Universal Robots URScript: Jonathan_code.script

  # Default parameters:
  global speed_ms = 0.3
  global speed_rads = 0.75
  global accel_mss = 3
  global accel_radss = 1.2
  global blend_radius_m = 0.001

  # Add subprograms here
  # Start of main program
  # Program generated by RoboDK v5.6.5 for UR10e on 12/10/2023 11:38:14
  # Using nominal kinematics.
  blend_radius_m = 0.001
  speed_ms = 1.000
  # set_reference(p[0.335000, -0.154000, 0.000000, 0.000000, 0.000000, 0.000000])
  set_tcp(p[0.000000, 0.000000, 0.253000, 0.000000, 0.000000, 0.000000])
  # Show Tool
  movej([0.470150, -1.112535, -2.574781, -1.025073, 1.570796, 2.040947],accel_radss,speed_rads,0,blend_radius_m
  movel([0.470150, -1.206188, -2.638649, -0.867552, 1.570796, 2.040947],accel_mss,speed_ms,0,blend_radius_m)
  speed_ms = 1.000
  movel([0.470150, -1.233460, -2.652834, -0.826095, 1.570796, 2.040947],accel_mss,speed_ms,0,blend_radius_m)
  speed_ms = 0.003
  movel([0.470150, -1.244207, -2.658024, -0.810158, 1.570796, 2.040947],accel_mss,speed_ms,0,blend_radius_m)
  speed_ms = 0.007
  movel([0.482800, -1.244203, -2.658026, -0.810160, 1.570796, 2.053597],accel_mss,speed_ms,0,blend_radius_m)
  movel([0.495365, -1.244373, -2.657937, -0.810079, 1.570796, 2.066162],accel_mss,speed_ms,0,blend_radius_m)
  movel([0.493680, -1.247797, -2.656131, -0.808461, 1.570796, 2.064476],accel_mss,speed_ms,0,blend_radius_m)
  movel([0.492007, -1.251200, -2.654322, -0.806866, 1.570796, 2.062803],accel_mss,speed_ms,0,blend_radius_m)
  movel([0.479519, -1.251033, -2.654411, -0.806944, 1.570796, 2.050316],accel_mss,speed_ms,0,blend_radius_m)
  movel([0.466949, -1.251037, -2.654410, -0.806943, 1.570796, 2.037745],accel_mss,speed_ms,0,blend_radius_m)
  movel([0.468544, -1.247632, -2.656219, -0.808539, 1.570796, 2.039340],accel_mss,speed_ms,0,blend_radius_m)
  movel([0.470150, -1.244207, -2.658024, -0.810158, 1.570796, 2.040947],accel_mss,speed_ms,0,blend_radius_m)
  speed_ms = 0.003
  movel([0.470150, -1.247853, -2.659738, -0.804798, 1.570796, 2.040947],accel_mss,speed_ms,0,blend_radius_m)
  speed_ms = 0.007
  movel([0.482800, -1.247850, -2.659740, -0.804799, 1.570796, 2.053597],accel_mss,speed_ms,0,blend_radius_m)
  movel([0.495365, -1.248020, -2.659650, -0.804719, 1.570796, 2.066162],accel_mss,speed_ms,0,blend_radius_m)
  movel([0.493680, -1.251437, -2.657839, -0.803114, 1.570796, 2.064476],accel_mss,speed_ms,0,blend_radius_m)
  movel([0.492007, -1.254834, -2.656024, -0.801531, 1.570796, 2.062803],accel_mss,speed_ms,0,blend_radius_m)
  movel([0.479519, -1.254667, -2.656113, -0.801608, 1.570796, 2.050316],accel_mss,speed_ms,0,blend_radius_m)
  movel([0.466949, -1.254671, -2.656111, -0.801607, 1.570796, 2.037745],accel_mss,speed_ms,0,blend_radius_m)
  movel([0.468544, -1.251272, -2.657926, -0.803191, 1.570796, 2.039340],accel_mss,speed_ms,0,blend_radius_m)
  movel([0.470150, -1.247853, -2.659738, -0.804798, 1.570796, 2.040947],accel_mss,speed_ms,0,blend_radius_m)
  speed_ms = 0.003
  movel([0.470150, -1.233460, -2.652834, -0.826095, 1.570796, 2.040947],accel_mss,speed_ms,0,blend_radius_m)
  speed_ms = 1.000
  movel([0.470150, -1.206188, -2.638649, -0.867552, 1.570796, 2.040947],accel_mss,speed_ms,0,blend_radius_m)
  movel([0.500005, -1.181387, -2.650684, -0.880318, 1.570796, 2.070801],accel_mss,speed_ms,0,blend_radius_m)
  movel([0.500005, -1.208894, -2.665198, -0.838297, 1.570796, 2.070801],accel_mss,speed_ms,0,blend_radius_m)
  speed_ms = 0.003
  movel([0.500005, -1.219758, -2.670513, -0.822118, 1.570796, 2.070801],accel_mss,speed_ms,0,blend_radius_m)
  speed_ms = 0.007
  movel([0.496713, -1.215452, -2.672641, -0.824296, 1.570796, 2.067509],accel_mss,speed_ms,0,blend_radius_m)
  movel([0.497565, -1.208277, -2.676141, -0.827971, 1.570796, 2.068361],accel_mss,speed_ms,0,blend_radius_m)
  movel([0.502312, -1.200573, -2.679835, -0.831981, 1.570796, 2.073109],accel_mss,speed_ms,0,blend_radius_m)
  movel([0.509447, -1.194948, -2.682491, -0.834950, 1.570796, 2.080243],accel_mss,speed_ms,0,blend_radius_m)
  movel([0.511019, -1.194268, -2.682810, -0.835312, 1.570796, 2.081816],accel_mss,speed_ms,0,blend_radius_m)
  movel([0.512848, -1.193698, -2.683076, -0.835615, 1.570796, 2.083644],accel_mss,speed_ms,0,blend_radius_m)
  movel([0.514636, -1.193318, -2.683254, -0.835817, 1.570796, 2.085432],accel_mss,speed_ms,0,blend_radius_m)
  movel([0.516087, -1.193207, -2.683306, -0.835876, 1.570796, 2.086884],accel_mss,speed_ms,0,blend_radius_m)
  movel([0.521675, -1.195790, -2.682095, -0.834503, 1.570796, 2.092471],accel_mss,speed_ms,0,blend_radius_m)
  movel([0.522729, -1.202299, -2.679013, -0.831077, 1.570796, 2.093526],accel_mss,speed_ms,0,blend_radius_m)
  movel([0.518940, -1.210348, -2.675137, -0.826904, 1.570796, 2.089737],accel_mss,speed_ms,0,blend_radius_m)
  movel([0.511727, -1.217078, -2.671840, -0.823471, 1.570796, 2.082524],accel_mss,speed_ms,0,blend_radius_m)
  movel([0.508244, -1.219012, -2.670883, -0.822493, 1.570796, 2.079040],accel_mss,speed_ms,0,blend_radius_m)
  movel([0.505130, -1.220107, -2.670340, -0.821942, 1.570796, 2.075926],accel_mss,speed_ms,0,blend_radius_m)
  movel([0.502386, -1.220345, -2.670222, -0.821823, 1.570796, 2.073182],accel_mss,speed_ms,0,blend_radius_m)
  movel([0.500005, -1.219758, -2.670513, -0.822118, 1.570796, 2.070801],accel_mss,speed_ms,0,blend_radius_m)
  speed_ms = 0.003
  movel([0.500005, -1.223447, -2.672269, -0.816673, 1.570796, 2.070801],accel_mss,speed_ms,0,blend_radius_m)
  speed_ms = 0.007
  movel([0.496713, -1.219148, -2.674405, -0.818836, 1.570796, 2.067509],accel_mss,speed_ms,0,blend_radius_m)
  movel([0.497565, -1.211984, -2.677917, -0.822488, 1.570796, 2.068361],accel_mss,speed_ms,0,blend_radius_m)
  movel([0.502312, -1.204292, -2.681624, -0.826473, 1.570796, 2.073109],accel_mss,speed_ms,0,blend_radius_m)
  movel([0.509447, -1.198675, -2.684289, -0.829425, 1.570796, 2.080243],accel_mss,speed_ms,0,blend_radius_m)
  movel([0.511019, -1.197995, -2.684609, -0.829784, 1.570796, 2.081816],accel_mss,speed_ms,0,blend_radius_m)
  movel([0.512848, -1.197426, -2.684877, -0.830086, 1.570796, 2.083644],accel_mss,speed_ms,0,blend_radius_m)
  movel([0.514636, -1.197048, -2.685055, -0.830287, 1.570796, 2.085432],accel_mss,speed_ms,0,blend_radius_m)
  movel([0.516087, -1.196936, -2.685107, -0.830346, 1.570796, 2.086884],accel_mss,speed_ms,0,blend_radius_m)
  movel([0.521675, -1.199516, -2.683892, -0.828981, 1.570796, 2.092471],accel_mss,speed_ms,0,blend_radius_m)
  movel([0.522729, -1.206015, -2.680799, -0.825575, 1.570796, 2.093526],accel_mss,speed_ms,0,blend_radius_m)
  movel([0.518940, -1.214052, -2.676909, -0.821428, 1.570796, 2.089737],accel_mss,speed_ms,0,blend_radius_m)
  movel([0.511727, -1.220771, -2.673601, -0.818017, 1.570796, 2.082524],accel_mss,speed_ms,0,blend_radius_m)
  movel([0.508244, -1.222703, -2.672640, -0.817046, 1.570796, 2.079040],accel_mss,speed_ms,0,blend_radius_m)
  movel([0.505130, -1.223795, -2.672095, -0.816499, 1.570796, 2.075926],accel_mss,speed_ms,0,blend_radius_m)
  movel([0.502386, -1.224033, -2.671976, -0.816380, 1.570796, 2.073182],accel_mss,speed_ms,0,blend_radius_m)
  movel([0.500005, -1.223447, -2.672269, -0.816673, 1.570796, 2.070801],accel_mss,speed_ms,0,blend_radius_m)
  speed_ms = 0.003
  movel([0.500005, -1.208894, -2.665198, -0.838297, 1.570796, 2.070801],accel_mss,speed_ms,0,blend_radius_m)
  speed_ms = 1.000
  movel([0.500005, -1.181387, -2.650684, -0.880318, 1.570796, 2.070801],accel_mss,speed_ms,0,blend_radius_m)
  movel([0.502939, -1.178463, -2.652060, -0.881866, 1.570796, 2.073735],accel_mss,speed_ms,0,blend_radius_m)
  movel([0.502939, -1.205994, -2.666612, -0.839782, 1.570796, 2.073735],accel_mss,speed_ms,0,blend_radius_m)
  speed_ms = 0.003
  movel([0.502939, -1.216871, -2.671942, -0.823575, 1.570796, 2.073735],accel_mss,speed_ms,0,blend_radius_m)
  speed_ms = 0.007
  movel([0.501818, -1.216382, -2.672184, -0.823824, 1.570796, 2.072614],accel_mss,speed_ms,0,blend_radius_m)
  movel([0.500967, -1.215437, -2.672649, -0.824303, 1.570796, 2.071763],accel_mss,speed_ms,0,blend_radius_m)
  movel([0.500167, -1.213807, -2.673449, -0.825133, 1.570796, 2.070964],accel_mss,speed_ms,0,blend_radius_m)
  movel([0.499493, -1.211784, -2.674438, -0.826167, 1.570796, 2.070289],accel_mss,speed_ms,0,blend_radius_m)
  movel([0.499454, -1.210389, -2.675117, -0.826883, 1.570796, 2.070250],accel_mss,speed_ms,0,blend_radius_m)
  movel([0.499992, -1.208799, -2.675888, -0.827701, 1.570796, 2.070788],accel_mss,speed_ms,0,blend_radius_m)
  movel([0.501476, -1.206040, -2.677221, -0.829128, 1.570796, 2.072272],accel_mss,speed_ms,0,blend_radius_m)
  movel([0.504659, -1.201513, -2.679388, -0.831488, 1.570796, 2.075455],accel_mss,speed_ms,0,blend_radius_m)
  movel([0.508226, -1.198314, -2.680906, -0.833169, 1.570796, 2.079022],accel_mss,speed_ms,0,blend_radius_m)
  movel([0.512021, -1.196627, -2.681702, -0.834060, 1.570796, 2.082817],accel_mss,speed_ms,0,blend_radius_m)
  movel([0.515863, -1.196480, -2.681771, -0.834138, 1.570796, 2.086659],accel_mss,speed_ms,0,blend_radius_m)
  movel([0.517050, -1.196870, -2.681587, -0.833932, 1.570796, 2.087846],accel_mss,speed_ms,0,blend_radius_m)
  movel([0.518044, -1.197576, -2.681254, -0.833558, 1.570796, 2.088840],accel_mss,speed_ms,0,blend_radius_m)
  movel([0.518815, -1.198576, -2.680782, -0.833031, 1.570796, 2.089612],accel_mss,speed_ms,0,blend_radius_m)
  movel([0.519336, -1.199836, -2.680185, -0.832368, 1.570796, 2.090133],accel_mss,speed_ms,0,blend_radius_m)
  movel([0.518927, -1.205179, -2.677634, -0.829575, 1.570796, 2.089724],accel_mss,speed_ms,0,blend_radius_m)
  movel([0.515430, -1.211016, -2.674812, -0.826561, 1.570796, 2.086227],accel_mss,speed_ms,0,blend_radius_m)
  movel([0.510067, -1.215433, -2.672651, -0.824305, 1.570796, 2.080863],accel_mss,speed_ms,0,blend_radius_m)
  movel([0.504562, -1.217042, -2.671858, -0.823489, 1.570796, 2.075358],accel_mss,speed_ms,0,blend_radius_m)
  movel([0.502939, -1.216871, -2.671942, -0.823575, 1.570796, 2.073735],accel_mss,speed_ms,0,blend_radius_m)
  speed_ms = 0.003
  movel([0.502939, -1.220565, -2.673703, -0.818121, 1.570796, 2.073735],accel_mss,speed_ms,0,blend_radius_m)
  speed_ms = 0.007
  movel([0.501818, -1.220076, -2.673945, -0.818367, 1.570796, 2.072614],accel_mss,speed_ms,0,blend_radius_m)
  movel([0.500967, -1.219134, -2.674412, -0.818844, 1.570796, 2.071763],accel_mss,speed_ms,0,blend_radius_m)
  movel([0.500167, -1.217506, -2.675215, -0.819668, 1.570796, 2.070964],accel_mss,speed_ms,0,blend_radius_m)
  movel([0.499493, -1.215486, -2.676207, -0.820696, 1.570796, 2.070289],accel_mss,speed_ms,0,blend_radius_m)
  movel([0.499454, -1.214093, -2.676889, -0.821407, 1.570796, 2.070250],accel_mss,speed_ms,0,blend_radius_m)
  movel([0.499992, -1.212506, -2.677663, -0.822220, 1.570796, 2.070788],accel_mss,speed_ms,0,blend_radius_m)
  movel([0.501476, -1.209751, -2.679000, -0.823638, 1.570796, 2.072272],accel_mss,speed_ms,0,blend_radius_m)
  movel([0.504659, -1.205231, -2.681175, -0.825983, 1.570796, 2.075455],accel_mss,speed_ms,0,blend_radius_m)
  movel([0.508226, -1.202036, -2.682698, -0.827655, 1.570796, 2.079022],accel_mss,speed_ms,0,blend_radius_m)
  movel([0.512021, -1.200352, -2.683497, -0.828540, 1.570796, 2.082817],accel_mss,speed_ms,0,blend_radius_m)
  movel([0.515863, -1.200205, -2.683566, -0.828617, 1.570796, 2.086659],accel_mss,speed_ms,0,blend_radius_m)
  movel([0.517050, -1.200594, -2.683382, -0.828413, 1.570796, 2.087846],accel_mss,speed_ms,0,blend_radius_m)
  movel([0.518044, -1.201300, -2.683048, -0.828041, 1.570796, 2.088840],accel_mss,speed_ms,0,blend_radius_m)
  movel([0.518815, -1.202298, -2.682574, -0.827517, 1.570796, 2.089612],accel_mss,speed_ms,0,blend_radius_m)
  movel([0.519336, -1.203556, -2.681975, -0.826858, 1.570796, 2.090133],accel_mss,speed_ms,0,blend_radius_m)
  movel([0.518927, -1.208892, -2.679415, -0.824082, 1.570796, 2.089724],accel_mss,speed_ms,0,blend_radius_m)
  movel([0.515430, -1.214719, -2.676583, -0.821087, 1.570796, 2.086227],accel_mss,speed_ms,0,blend_radius_m)
  movel([0.510067, -1.219129, -2.674414, -0.818846, 1.570796, 2.080863],accel_mss,speed_ms,0,blend_radius_m)
  movel([0.504562, -1.220735, -2.673619, -0.818035, 1.570796, 2.075358],accel_mss,speed_ms,0,blend_radius_m)
  movel([0.502939, -1.220565, -2.673703, -0.818121, 1.570796, 2.073735],accel_mss,speed_ms,0,blend_radius_m)
  speed_ms = 0.003
  movel([0.502939, -1.205994, -2.666612, -0.839782, 1.570796, 2.073735],accel_mss,speed_ms,0,blend_radius_m)
  speed_ms = 1.000
  movel([0.502939, -1.178463, -2.652060, -0.881866, 1.570796, 2.073735],accel_mss,speed_ms,0,blend_radius_m)
  movel([0.506130, -1.175000, -2.653677, -0.883712, 1.570796, 2.076926],accel_mss,speed_ms,0,blend_radius_m)
  movel([0.506130, -1.202560, -2.668276, -0.841553, 1.570796, 2.076926],accel_mss,speed_ms,0,blend_radius_m)
  speed_ms = 0.003
  movel([0.506130, -1.213452, -2.673623, -0.825314, 1.570796, 2.076926],accel_mss,speed_ms,0,blend_radius_m)
  speed_ms = 0.007
  movel([0.503262, -1.211890, -2.674386, -0.826113, 1.570796, 2.074059],accel_mss,speed_ms,0,blend_radius_m)
  movel([0.503107, -1.207977, -2.676286, -0.828126, 1.570796, 2.073904],accel_mss,speed_ms,0,blend_radius_m)
  movel([0.505736, -1.203530, -2.678425, -0.830434, 1.570796, 2.076532],accel_mss,speed_ms,0,blend_radius_m)
  movel([0.509953, -1.200615, -2.679815, -0.831959, 1.570796, 2.080749],accel_mss,speed_ms,0,blend_radius_m)
  movel([0.512348, -1.199943, -2.680134, -0.832312, 1.570796, 2.083144],accel_mss,speed_ms,0,blend_radius_m)
  movel([0.514007, -1.199944, -2.680134, -0.832311, 1.570796, 2.084803],accel_mss,speed_ms,0,blend_radius_m)
  movel([0.515159, -1.200632, -2.679807, -0.831950, 1.570796, 2.085955],accel_mss,speed_ms,0,blend_radius_m)
  movel([0.515994, -1.202071, -2.679122, -0.831196, 1.570796, 2.086790],accel_mss,speed_ms,0,blend_radius_m)
  movel([0.515943, -1.205637, -2.677415, -0.829338, 1.570796, 2.086739],accel_mss,speed_ms,0,blend_radius_m)
  movel([0.513721, -1.209501, -2.675548, -0.827340, 1.570796, 2.084517],accel_mss,speed_ms,0,blend_radius_m)
  movel([0.510054, -1.212409, -2.674133, -0.825847, 1.570796, 2.080851],accel_mss,speed_ms,0,blend_radius_m)
  movel([0.506130, -1.213452, -2.673623, -0.825314, 1.570796, 2.076926],accel_mss,speed_ms,0,blend_radius_m)
  speed_ms = 0.003
  movel([0.506130, -1.217151, -2.675389, -0.819848, 1.570796, 2.076926],accel_mss,speed_ms,0,blend_radius_m)
  speed_ms = 0.007
  movel([0.503262, -1.215592, -2.676155, -0.820642, 1.570796, 2.074059],accel_mss,speed_ms,0,blend_radius_m)
  movel([0.503107, -1.211685, -2.678062, -0.822642, 1.570796, 2.073904],accel_mss,speed_ms,0,blend_radius_m)
  movel([0.505736, -1.207244, -2.680209, -0.824936, 1.570796, 2.076532],accel_mss,speed_ms,0,blend_radius_m)
  movel([0.509953, -1.204334, -2.681603, -0.826451, 1.570796, 2.080749],accel_mss,speed_ms,0,blend_radius_m)
  movel([0.512348, -1.203663, -2.681924, -0.826802, 1.570796, 2.083144],accel_mss,speed_ms,0,blend_radius_m)
  movel([0.514007, -1.203664, -2.681924, -0.826802, 1.570796, 2.084803],accel_mss,speed_ms,0,blend_radius_m)
  movel([0.515159, -1.204351, -2.681596, -0.826443, 1.570796, 2.085955],accel_mss,speed_ms,0,blend_radius_m)
  movel([0.515994, -1.205787, -2.680908, -0.825693, 1.570796, 2.086790],accel_mss,speed_ms,0,blend_radius_m)
  movel([0.515943, -1.209348, -2.679194, -0.823846, 1.570796, 2.086739],accel_mss,speed_ms,0,blend_radius_m)
  movel([0.513721, -1.213207, -2.677321, -0.821861, 1.570796, 2.084517],accel_mss,speed_ms,0,blend_radius_m)
  movel([0.510054, -1.216110, -2.675901, -0.820378, 1.570796, 2.080851],accel_mss,speed_ms,0,blend_radius_m)
  movel([0.506130, -1.217151, -2.675389, -0.819848, 1.570796, 2.076926],accel_mss,speed_ms,0,blend_radius_m)
  speed_ms = 0.003
  movel([0.506130, -1.202560, -2.668276, -0.841553, 1.570796, 2.076926],accel_mss,speed_ms,0,blend_radius_m)
  speed_ms = 1.000
  movel([0.506130, -1.175000, -2.653677, -0.883712, 1.570796, 2.076926],accel_mss,speed_ms,0,blend_radius_m)
  movel([0.511926, -1.148900, -2.665470, -0.898018, 1.570796, 2.082723],accel_mss,speed_ms,0,blend_radius_m)
  movel([0.511926, -1.176644, -2.680413, -0.855332, 1.570796, 2.082723],accel_mss,speed_ms,0,blend_radius_m)
  speed_ms = 0.003
  movel([0.511926, -1.187635, -2.685892, -0.838862, 1.570796, 2.082723],accel_mss,speed_ms,0,blend_radius_m)
  speed_ms = 0.007
  movel([0.498596, -1.192917, -2.683441, -0.836031, 1.570796, 2.069392],accel_mss,speed_ms,0,blend_radius_m)
  movel([0.503810, -1.182117, -2.688420, -0.841852, 1.570796, 2.074606],accel_mss,speed_ms,0,blend_radius_m)
  movel([0.509142, -1.171113, -2.693365, -0.847911, 1.570796, 2.079938],accel_mss,speed_ms,0,blend_radius_m)
  movel([0.511240, -1.172435, -2.692778, -0.847176, 1.570796, 2.082036],accel_mss,speed_ms,0,blend_radius_m)
  movel([0.517671, -1.176577, -2.690926, -0.844886, 1.570796, 2.088468],accel_mss,speed_ms,0,blend_radius_m)
  movel([0.521715, -1.179304, -2.689697, -0.843389, 1.570796, 2.092511],accel_mss,speed_ms,0,blend_radius_m)
  movel([0.524550, -1.181302, -2.688791, -0.842296, 1.570796, 2.095346],accel_mss,speed_ms,0,blend_radius_m)
  movel([0.525020, -1.181849, -2.688542, -0.841998, 1.570796, 2.095816],accel_mss,speed_ms,0,blend_radius_m)
  movel([0.524802, -1.182217, -2.688375, -0.841797, 1.570796, 2.095598],accel_mss,speed_ms,0,blend_radius_m)
  movel([0.521291, -1.183784, -2.687660, -0.840945, 1.570796, 2.092088],accel_mss,speed_ms,0,blend_radius_m)
  movel([0.517034, -1.185590, -2.686833, -0.839966, 1.570796, 2.087830],accel_mss,speed_ms,0,blend_radius_m)
  movel([0.511926, -1.187635, -2.685892, -0.838862, 1.570796, 2.082723],accel_mss,speed_ms,0,blend_radius_m)
  speed_ms = 0.003
  movel([0.511926, -1.191372, -2.687703, -0.833314, 1.570796, 2.082723],accel_mss,speed_ms,0,blend_radius_m)
  speed_ms = 0.007
  movel([0.498596, -1.196647, -2.685243, -0.830499, 1.570796, 2.069392],accel_mss,speed_ms,0,blend_radius_m)
  movel([0.503810, -1.185861, -2.690240, -0.836288, 1.570796, 2.074606],accel_mss,speed_ms,0,blend_radius_m)
  movel([0.509142, -1.174870, -2.695204, -0.842315, 1.570796, 2.079938],accel_mss,speed_ms,0,blend_radius_m)
  movel([0.511240, -1.176191, -2.694614, -0.841584, 1.570796, 2.082036],accel_mss,speed_ms,0,blend_radius_m)
  movel([0.517671, -1.180327, -2.692755, -0.839306, 1.570796, 2.088468],accel_mss,speed_ms,0,blend_radius_m)
  movel([0.521715, -1.183051, -2.691522, -0.837816, 1.570796, 2.092511],accel_mss,speed_ms,0,blend_radius_m)
  movel([0.524550, -1.185047, -2.690612, -0.836730, 1.570796, 2.095346],accel_mss,speed_ms,0,blend_radius_m)
  movel([0.525020, -1.185593, -2.690363, -0.836433, 1.570796, 2.095816],accel_mss,speed_ms,0,blend_radius_m)
  movel([0.524802, -1.185961, -2.690195, -0.836234, 1.570796, 2.095598],accel_mss,speed_ms,0,blend_radius_m)
  movel([0.521291, -1.187526, -2.689477, -0.835386, 1.570796, 2.092088],accel_mss,speed_ms,0,blend_radius_m)
  movel([0.517034, -1.189329, -2.688647, -0.834413, 1.570796, 2.087830],accel_mss,speed_ms,0,blend_radius_m)
  movel([0.511926, -1.191372, -2.687703, -0.833314, 1.570796, 2.082723],accel_mss,speed_ms,0,blend_radius_m)
  speed_ms = 0.003
  movel([0.511926, -1.176644, -2.680413, -0.855332, 1.570796, 2.082723],accel_mss,speed_ms,0,blend_radius_m)
  speed_ms = 1.000
  movel([0.511926, -1.148900, -2.665470, -0.898018, 1.570796, 2.082723],accel_mss,speed_ms,0,blend_radius_m)
  movel([0.484054, -1.150700, -2.664679, -0.897010, 1.570796, 2.054851],accel_mss,speed_ms,0,blend_radius_m)
  movel([0.484054, -1.178433, -2.679598, -0.854358, 1.570796, 2.054851],accel_mss,speed_ms,0,blend_radius_m)
  speed_ms = 0.003
  movel([0.484054, -1.189418, -2.685068, -0.837903, 1.570796, 2.054851],accel_mss,speed_ms,0,blend_radius_m)
  speed_ms = 0.007
  movel([0.480506, -1.198853, -2.680651, -0.832885, 1.570796, 2.051303],accel_mss,speed_ms,0,blend_radius_m)
  movel([0.477443, -1.208248, -2.676155, -0.827986, 1.570796, 2.048239],accel_mss,speed_ms,0,blend_radius_m)
  movel([0.476365, -1.210715, -2.674959, -0.826715, 1.570796, 2.047161],accel_mss,speed_ms,0,blend_radius_m)
  movel([0.475147, -1.211860, -2.674401, -0.826128, 1.570796, 2.045943],accel_mss,speed_ms,0,blend_radius_m)
  movel([0.473142, -1.212453, -2.674111, -0.825825, 1.570796, 2.043939],accel_mss,speed_ms,0,blend_radius_m)
  movel([0.471647, -1.212536, -2.674071, -0.825782, 1.570796, 2.042444],accel_mss,speed_ms,0,blend_radius_m)
  movel([0.470897, -1.212281, -2.674195, -0.825912, 1.570796, 2.041693],accel_mss,speed_ms,0,blend_radius_m)
  movel([0.470592, -1.211613, -2.674521, -0.826255, 1.570796, 2.041389],accel_mss,speed_ms,0,blend_radius_m)
  movel([0.470632, -1.210285, -2.675167, -0.826936, 1.570796, 2.041428],accel_mss,speed_ms,0,blend_radius_m)
  movel([0.473573, -1.198109, -2.681003, -0.833277, 1.570796, 2.044369],accel_mss,speed_ms,0,blend_radius_m)
  movel([0.480363, -1.181578, -2.688665, -0.842146, 1.570796, 2.051160],accel_mss,speed_ms,0,blend_radius_m)
  movel([0.489208, -1.164498, -2.696277, -0.851614, 1.570796, 2.060004],accel_mss,speed_ms,0,blend_radius_m)
  movel([0.498310, -1.151098, -2.702038, -0.859253, 1.570796, 2.069106],accel_mss,speed_ms,0,blend_radius_m)
  movel([0.499374, -1.149933, -2.702530, -0.859926, 1.570796, 2.070170],accel_mss,speed_ms,0,blend_radius_m)
  movel([0.500392, -1.149174, -2.702850, -0.860365, 1.570796, 2.071188],accel_mss,speed_ms,0,blend_radius_m)
  movel([0.501497, -1.148747, -2.703030, -0.860612, 1.570796, 2.072293],accel_mss,speed_ms,0,blend_radius_m)
  movel([0.502836, -1.148585, -2.703098, -0.860706, 1.570796, 2.073632],accel_mss,speed_ms,0,blend_radius_m)
  movel([0.503826, -1.148619, -2.703084, -0.860686, 1.570796, 2.074623],accel_mss,speed_ms,0,blend_radius_m)
  movel([0.504671, -1.148774, -2.703018, -0.860597, 1.570796, 2.075467],accel_mss,speed_ms,0,blend_radius_m)
  movel([0.505282, -1.149008, -2.702920, -0.860461, 1.570796, 2.076078],accel_mss,speed_ms,0,blend_radius_m)
  movel([0.505458, -1.149307, -2.702794, -0.860288, 1.570796, 2.076254],accel_mss,speed_ms,0,blend_radius_m)
  movel([0.505300, -1.149879, -2.702553, -0.859957, 1.570796, 2.076096],accel_mss,speed_ms,0,blend_radius_m)
  movel([0.504211, -1.151773, -2.701752, -0.858864, 1.570796, 2.075007],accel_mss,speed_ms,0,blend_radius_m)
  movel([0.502820, -1.154048, -2.700785, -0.857556, 1.570796, 2.073616],accel_mss,speed_ms,0,blend_radius_m)
  movel([0.501171, -1.156589, -2.699699, -0.856101, 1.570796, 2.071967],accel_mss,speed_ms,0,blend_radius_m)
  movel([0.495509, -1.165940, -2.695646, -0.850803, 1.570796, 2.066305],accel_mss,speed_ms,0,blend_radius_m)
  movel([0.489418, -1.177710, -2.690416, -0.844263, 1.570796, 2.060214],accel_mss,speed_ms,0,blend_radius_m)
  movel([0.484054, -1.189418, -2.685068, -0.837903, 1.570796, 2.054851],accel_mss,speed_ms,0,blend_radius_m)
  speed_ms = 0.003
  movel([0.484054, -1.193152, -2.686876, -0.832361, 1.570796, 2.054851],accel_mss,speed_ms,0,blend_radius_m)
  speed_ms = 0.007
  movel([0.480506, -1.202575, -2.682442, -0.827372, 1.570796, 2.051303],accel_mss,speed_ms,0,blend_radius_m)
  movel([0.477443, -1.211956, -2.677931, -0.822503, 1.570796, 2.048239],accel_mss,speed_ms,0,blend_radius_m)
  movel([0.476365, -1.214419, -2.676730, -0.821241, 1.570796, 2.047161],accel_mss,speed_ms,0,blend_radius_m)
  movel([0.475147, -1.215562, -2.676170, -0.820657, 1.570796, 2.045943],accel_mss,speed_ms,0,blend_radius_m)
  movel([0.473142, -1.216154, -2.675879, -0.820355, 1.570796, 2.043939],accel_mss,speed_ms,0,blend_radius_m)
  movel([0.471647, -1.216237, -2.675839, -0.820313, 1.570796, 2.042444],accel_mss,speed_ms,0,blend_radius_m)
  movel([0.470897, -1.215983, -2.675964, -0.820443, 1.570796, 2.041693],accel_mss,speed_ms,0,blend_radius_m)
  movel([0.470592, -1.215315, -2.676291, -0.820783, 1.570796, 2.041389],accel_mss,speed_ms,0,blend_radius_m)
  movel([0.470632, -1.213990, -2.676939, -0.821460, 1.570796, 2.041428],accel_mss,speed_ms,0,blend_radius_m)
  movel([0.473573, -1.201831, -2.682796, -0.827762, 1.570796, 2.044369],accel_mss,speed_ms,0,blend_radius_m)
  movel([0.480363, -1.185322, -2.690487, -0.836580, 1.570796, 2.051160],accel_mss,speed_ms,0,blend_radius_m)
  movel([0.489208, -1.168263, -2.698127, -0.845999, 1.570796, 2.060004],accel_mss,speed_ms,0,blend_radius_m)
  movel([0.498310, -1.154875, -2.703911, -0.853603, 1.570796, 2.069106],accel_mss,speed_ms,0,blend_radius_m)
  movel([0.499374, -1.153712, -2.704405, -0.854272, 1.570796, 2.070170],accel_mss,speed_ms,0,blend_radius_m)
  movel([0.500392, -1.152953, -2.704726, -0.854710, 1.570796, 2.071188],accel_mss,speed_ms,0,blend_radius_m)
  movel([0.501497, -1.152526, -2.704907, -0.854956, 1.570796, 2.072293],accel_mss,speed_ms,0,blend_radius_m)
  movel([0.502836, -1.152365, -2.704975, -0.855049, 1.570796, 2.073632],accel_mss,speed_ms,0,blend_radius_m)
  movel([0.503826, -1.152398, -2.704961, -0.855030, 1.570796, 2.074623],accel_mss,speed_ms,0,blend_radius_m)
  movel([0.504671, -1.152553, -2.704895, -0.854940, 1.570796, 2.075467],accel_mss,speed_ms,0,blend_radius_m)
  movel([0.505282, -1.152787, -2.704797, -0.854806, 1.570796, 2.076078],accel_mss,speed_ms,0,blend_radius_m)
  movel([0.505458, -1.153086, -2.704670, -0.854633, 1.570796, 2.076254],accel_mss,speed_ms,0,blend_radius_m)
  movel([0.505300, -1.153657, -2.704428, -0.854304, 1.570796, 2.076096],accel_mss,speed_ms,0,blend_radius_m)
  movel([0.504211, -1.155550, -2.703624, -0.853215, 1.570796, 2.075007],accel_mss,speed_ms,0,blend_radius_m)
  movel([0.502820, -1.157822, -2.702653, -0.851913, 1.570796, 2.073616],accel_mss,speed_ms,0,blend_radius_m)
  movel([0.501171, -1.160361, -2.701563, -0.850465, 1.570796, 2.071967],accel_mss,speed_ms,0,blend_radius_m)
  movel([0.495509, -1.169702, -2.697494, -0.845192, 1.570796, 2.066305],accel_mss,speed_ms,0,blend_radius_m)
  movel([0.489418, -1.181459, -2.692244, -0.838686, 1.570796, 2.060214],accel_mss,speed_ms,0,blend_radius_m)
  movel([0.484054, -1.193152, -2.686876, -0.832361, 1.570796, 2.054851],accel_mss,speed_ms,0,blend_radius_m)
  speed_ms = 0.003
  movel([0.484054, -1.178433, -2.679598, -0.854358, 1.570796, 2.054851],accel_mss,speed_ms,0,blend_radius_m)
  speed_ms = 1.000
  movel([0.484054, -1.150700, -2.664679, -0.897010, 1.570796, 2.054851],accel_mss,speed_ms,0,blend_radius_m)
  movel([0.523020, -1.125862, -2.675313, -0.911214, 1.570796, 2.093816],accel_mss,speed_ms,0,blend_radius_m)
  movel([0.523020, -1.153722, -2.690557, -0.868110, 1.570796, 2.093816],accel_mss,speed_ms,0,blend_radius_m)
  speed_ms = 0.003
  movel([0.523020, -1.164783, -2.696152, -0.851453, 1.570796, 2.093816],accel_mss,speed_ms,0,blend_radius_m)
  speed_ms = 0.007
  movel([0.522684, -1.157268, -2.699408, -0.855713, 1.570796, 2.093481],accel_mss,speed_ms,0,blend_radius_m)
  movel([0.524949, -1.152033, -2.701642, -0.858714, 1.570796, 2.095745],accel_mss,speed_ms,0,blend_radius_m)
  movel([0.528948, -1.146645, -2.703912, -0.861832, 1.570796, 2.099745],accel_mss,speed_ms,0,blend_radius_m)
  movel([0.533936, -1.142070, -2.705817, -0.864502, 1.570796, 2.104732],accel_mss,speed_ms,0,blend_radius_m)
  movel([0.539020, -1.139206, -2.706999, -0.866184, 1.570796, 2.109816],accel_mss,speed_ms,0,blend_radius_m)
  movel([0.546147, -1.138732, -2.707194, -0.866463, 1.570796, 2.116944],accel_mss,speed_ms,0,blend_radius_m)
  movel([0.549993, -1.143138, -2.705374, -0.863877, 1.570796, 2.120789],accel_mss,speed_ms,0,blend_radius_m)
  movel([0.549294, -1.150892, -2.702125, -0.859372, 1.570796, 2.120091],accel_mss,speed_ms,0,blend_radius_m)
  movel([0.544338, -1.159300, -2.698534, -0.854555, 1.570796, 2.115134],accel_mss,speed_ms,0,blend_radius_m)
  movel([0.536255, -1.166000, -2.695620, -0.850769, 1.570796, 2.107051],accel_mss,speed_ms,0,blend_radius_m)
  movel([0.528182, -1.168073, -2.694709, -0.849607, 1.570796, 2.098978],accel_mss,speed_ms,0,blend_radius_m)
  movel([0.523020, -1.164783, -2.696152, -0.851453, 1.570796, 2.093816],accel_mss,speed_ms,0,blend_radius_m)
  speed_ms = 0.003
  movel([0.523020, -1.168547, -2.698002, -0.845840, 1.570796, 2.093816],accel_mss,speed_ms,0,blend_radius_m)
  speed_ms = 0.007
  movel([0.522684, -1.161039, -2.701271, -0.850079, 1.570796, 2.093481],accel_mss,speed_ms,0,blend_radius_m)
  movel([0.524949, -1.155809, -2.703513, -0.853066, 1.570796, 2.095745],accel_mss,speed_ms,0,blend_radius_m)
  movel([0.528948, -1.150427, -2.705792, -0.856170, 1.570796, 2.099745],accel_mss,speed_ms,0,blend_radius_m)
  movel([0.533936, -1.145855, -2.707705, -0.858829, 1.570796, 2.104732],accel_mss,speed_ms,0,blend_radius_m)
  movel([0.539020, -1.142993, -2.708892, -0.860504, 1.570796, 2.109816],accel_mss,speed_ms,0,blend_radius_m)
  movel([0.546147, -1.142519, -2.709087, -0.860782, 1.570796, 2.116944],accel_mss,speed_ms,0,blend_radius_m)
  movel([0.549993, -1.146923, -2.707260, -0.858206, 1.570796, 2.120789],accel_mss,speed_ms,0,blend_radius_m)
  movel([0.549294, -1.154669, -2.703998, -0.853721, 1.570796, 2.120091],accel_mss,speed_ms,0,blend_radius_m)
  movel([0.544338, -1.163069, -2.700393, -0.848927, 1.570796, 2.115134],accel_mss,speed_ms,0,blend_radius_m)
  movel([0.536255, -1.169762, -2.697468, -0.845159, 1.570796, 2.107051],accel_mss,speed_ms,0,blend_radius_m)
  movel([0.528182, -1.171833, -2.696553, -0.844002, 1.570796, 2.098978],accel_mss,speed_ms,0,blend_radius_m)
  movel([0.523020, -1.168547, -2.698002, -0.845840, 1.570796, 2.093816],accel_mss,speed_ms,0,blend_radius_m)
  speed_ms = 0.003
  movel([0.523020, -1.153722, -2.690557, -0.868110, 1.570796, 2.093816],accel_mss,speed_ms,0,blend_radius_m)
  speed_ms = 1.000
  movel([0.523020, -1.125862, -2.675313, -0.911214, 1.570796, 2.093816],accel_mss,speed_ms,0,blend_radius_m)
  movel([0.525596, -1.120968, -2.677337, -0.914083, 1.570796, 2.096393],accel_mss,speed_ms,0,blend_radius_m)
  movel([0.525596, -1.148847, -2.692645, -0.870896, 1.570796, 2.096393],accel_mss,speed_ms,0,blend_radius_m)
  speed_ms = 0.003
  movel([0.525596, -1.159922, -2.698265, -0.854202, 1.570796, 2.096393],accel_mss,speed_ms,0,blend_radius_m)
  speed_ms = 0.007
  movel([0.527217, -1.153485, -2.701025, -0.857879, 1.570796, 2.098013],accel_mss,speed_ms,0,blend_radius_m)
  movel([0.531860, -1.146983, -2.703770, -0.861636, 1.570796, 2.102656],accel_mss,speed_ms,0,blend_radius_m)
  movel([0.537911, -1.142814, -2.705508, -0.864066, 1.570796, 2.108707],accel_mss,speed_ms,0,blend_radius_m)
  movel([0.540711, -1.141772, -2.705940, -0.864677, 1.570796, 2.111507],accel_mss,speed_ms,0,blend_radius_m)
  movel([0.542057, -1.141528, -2.706041, -0.864820, 1.570796, 2.112854],accel_mss,speed_ms,0,blend_radius_m)
  movel([0.543149, -1.141793, -2.705931, -0.864664, 1.570796, 2.113946],accel_mss,speed_ms,0,blend_radius_m)
  movel([0.544875, -1.142872, -2.705485, -0.864033, 1.570796, 2.115671],accel_mss,speed_ms,0,blend_radius_m)
  movel([0.546522, -1.144687, -2.704730, -0.862972, 1.570796, 2.117319],accel_mss,speed_ms,0,blend_radius_m)
  movel([0.547091, -1.147035, -2.703748, -0.861605, 1.570796, 2.117887],accel_mss,speed_ms,0,blend_radius_m)
  movel([0.546568, -1.150041, -2.702484, -0.859863, 1.570796, 2.117365],accel_mss,speed_ms,0,blend_radius_m)
  movel([0.544975, -1.153815, -2.700885, -0.857690, 1.570796, 2.115771],accel_mss,speed_ms,0,blend_radius_m)
  movel([0.541190, -1.159267, -2.698548, -0.854574, 1.570796, 2.111986],accel_mss,speed_ms,0,blend_radius_m)
  movel([0.536401, -1.163211, -2.696838, -0.852339, 1.570796, 2.107198],accel_mss,speed_ms,0,blend_radius_m)
  movel([0.531558, -1.164876, -2.696112, -0.851401, 1.570796, 2.102354],accel_mss,speed_ms,0,blend_radius_m)
  movel([0.527584, -1.164010, -2.696490, -0.851889, 1.570796, 2.098380],accel_mss,speed_ms,0,blend_radius_m)
  movel([0.525596, -1.159922, -2.698265, -0.854202, 1.570796, 2.096393],accel_mss,speed_ms,0,blend_radius_m)
  speed_ms = 0.003
  movel([0.525596, -1.163691, -2.700123, -0.848575, 1.570796, 2.096393],accel_mss,speed_ms,0,blend_radius_m)
  speed_ms = 0.007
  movel([0.527217, -1.157260, -2.702894, -0.852235, 1.570796, 2.098013],accel_mss,speed_ms,0,blend_radius_m)
  movel([0.531860, -1.150764, -2.705650, -0.855975, 1.570796, 2.102656],accel_mss,speed_ms,0,blend_radius_m)
  movel([0.537911, -1.146599, -2.707395, -0.858395, 1.570796, 2.108707],accel_mss,speed_ms,0,blend_radius_m)
  movel([0.540711, -1.145557, -2.707829, -0.859003, 1.570796, 2.111507],accel_mss,speed_ms,0,blend_radius_m)
  movel([0.542057, -1.145313, -2.707930, -0.859145, 1.570796, 2.112854],accel_mss,speed_ms,0,blend_radius_m)
  movel([0.543149, -1.145578, -2.707820, -0.858990, 1.570796, 2.113946],accel_mss,speed_ms,0,blend_radius_m)
  movel([0.544875, -1.146656, -2.707371, -0.858362, 1.570796, 2.115671],accel_mss,speed_ms,0,blend_radius_m)
  movel([0.546522, -1.148470, -2.706614, -0.857306, 1.570796, 2.117319],accel_mss,speed_ms,0,blend_radius_m)
  movel([0.547091, -1.150816, -2.705628, -0.855945, 1.570796, 2.117887],accel_mss,speed_ms,0,blend_radius_m)
  movel([0.546568, -1.153820, -2.704359, -0.854210, 1.570796, 2.117365],accel_mss,speed_ms,0,blend_radius_m)
  movel([0.544975, -1.157589, -2.702753, -0.852047, 1.570796, 2.115771],accel_mss,speed_ms,0,blend_radius_m)
  movel([0.541190, -1.163037, -2.700407, -0.848945, 1.570796, 2.111986],accel_mss,speed_ms,0,blend_radius_m)
  movel([0.536401, -1.166977, -2.698691, -0.846722, 1.570796, 2.107198],accel_mss,speed_ms,0,blend_radius_m)
  movel([0.531558, -1.168640, -2.697962, -0.845788, 1.570796, 2.102354],accel_mss,speed_ms,0,blend_radius_m)
  movel([0.527584, -1.167774, -2.698341, -0.846273, 1.570796, 2.098380],accel_mss,speed_ms,0,blend_radius_m)
  movel([0.525596, -1.163691, -2.700123, -0.848575, 1.570796, 2.096393],accel_mss,speed_ms,0,blend_radius_m)
  speed_ms = 0.003
  movel([0.525596, -1.148847, -2.692645, -0.870896, 1.570796, 2.096393],accel_mss,speed_ms,0,blend_radius_m)
  speed_ms = 1.000
  movel([0.525596, -1.120968, -2.677337, -0.914083, 1.570796, 2.096393],accel_mss,speed_ms,0,blend_radius_m)
  movel([0.529262, -1.117192, -2.678884, -0.916313, 1.570796, 2.100059],accel_mss,speed_ms,0,blend_radius_m)
  movel([0.529262, -1.145084, -2.694241, -0.873064, 1.570796, 2.100059],accel_mss,speed_ms,0,blend_radius_m)
  speed_ms = 0.003
  movel([0.529262, -1.156168, -2.699880, -0.856341, 1.570796, 2.100059],accel_mss,speed_ms,0,blend_radius_m)
  speed_ms = 0.007
  movel([0.529392, -1.154530, -2.700580, -0.857279, 1.570796, 2.100188],accel_mss,speed_ms,0,blend_radius_m)
  movel([0.529749, -1.153424, -2.701051, -0.857914, 1.570796, 2.100545],accel_mss,speed_ms,0,blend_radius_m)
  movel([0.530494, -1.152320, -2.701520, -0.858549, 1.570796, 2.101290],accel_mss,speed_ms,0,blend_radius_m)
  movel([0.531998, -1.150687, -2.702211, -0.859490, 1.570796, 2.102795],accel_mss,speed_ms,0,blend_radius_m)
  movel([0.533218, -1.149554, -2.702690, -0.860145, 1.570796, 2.104014],accel_mss,speed_ms,0,blend_radius_m)
  movel([0.534676, -1.148406, -2.703173, -0.860810, 1.570796, 2.105473],accel_mss,speed_ms,0,blend_radius_m)
  movel([0.536130, -1.147419, -2.703588, -0.861383, 1.570796, 2.106926],accel_mss,speed_ms,0,blend_radius_m)
  movel([0.537342, -1.146768, -2.703861, -0.861761, 1.570796, 2.108138],accel_mss,speed_ms,0,blend_radius_m)
  movel([0.540988, -1.146278, -2.704066, -0.862046, 1.570796, 2.111785],accel_mss,speed_ms,0,blend_radius_m)
  movel([0.543117, -1.148292, -2.703221, -0.860876, 1.570796, 2.113913],accel_mss,speed_ms,0,blend_radius_m)
  movel([0.542994, -1.152091, -2.701617, -0.858681, 1.570796, 2.113790],accel_mss,speed_ms,0,blend_radius_m)
  movel([0.540654, -1.156319, -2.699815, -0.856255, 1.570796, 2.111450],accel_mss,speed_ms,0,blend_radius_m)
  movel([0.536970, -1.159496, -2.698449, -0.854444, 1.570796, 2.107766],accel_mss,speed_ms,0,blend_radius_m)
  movel([0.533123, -1.160663, -2.697944, -0.853781, 1.570796, 2.103919],accel_mss,speed_ms,0,blend_radius_m)
  movel([0.530256, -1.159437, -2.698475, -0.854478, 1.570796, 2.101052],accel_mss,speed_ms,0,blend_radius_m)
  movel([0.529262, -1.156168, -2.699880, -0.856341, 1.570796, 2.100059],accel_mss,speed_ms,0,blend_radius_m)
  speed_ms = 0.003
  movel([0.529262, -1.159941, -2.701744, -0.850704, 1.570796, 2.100059],accel_mss,speed_ms,0,blend_radius_m)
  speed_ms = 0.007
  movel([0.529392, -1.158304, -2.702447, -0.851638, 1.570796, 2.100188],accel_mss,speed_ms,0,blend_radius_m)
  movel([0.529749, -1.157199, -2.702920, -0.852270, 1.570796, 2.100545],accel_mss,speed_ms,0,blend_radius_m)
  movel([0.530494, -1.156097, -2.703391, -0.852902, 1.570796, 2.101290],accel_mss,speed_ms,0,blend_radius_m)
  movel([0.531998, -1.154465, -2.704085, -0.853839, 1.570796, 2.102795],accel_mss,speed_ms,0,blend_radius_m)
  movel([0.533218, -1.153333, -2.704565, -0.854491, 1.570796, 2.104014],accel_mss,speed_ms,0,blend_radius_m)
  movel([0.534676, -1.152185, -2.705051, -0.855153, 1.570796, 2.105473],accel_mss,speed_ms,0,blend_radius_m)
  movel([0.536130, -1.151199, -2.705467, -0.855723, 1.570796, 2.106926],accel_mss,speed_ms,0,blend_radius_m)
  movel([0.537342, -1.150549, -2.705741, -0.856099, 1.570796, 2.108138],accel_mss,speed_ms,0,blend_radius_m)
  movel([0.540988, -1.150059, -2.705947, -0.856383, 1.570796, 2.111785],accel_mss,speed_ms,0,blend_radius_m)
  movel([0.543117, -1.152071, -2.705099, -0.855219, 1.570796, 2.113913],accel_mss,speed_ms,0,blend_radius_m)
  movel([0.542994, -1.155867, -2.703489, -0.853033, 1.570796, 2.113790],accel_mss,speed_ms,0,blend_radius_m)
  movel([0.540654, -1.160091, -2.701679, -0.850619, 1.570796, 2.111450],accel_mss,speed_ms,0,blend_radius_m)
  movel([0.536970, -1.163265, -2.700308, -0.848816, 1.570796, 2.107766],accel_mss,speed_ms,0,blend_radius_m)
  movel([0.533123, -1.164431, -2.699801, -0.848157, 1.570796, 2.103919],accel_mss,speed_ms,0,blend_radius_m)
  movel([0.530256, -1.163206, -2.700333, -0.848850, 1.570796, 2.101052],accel_mss,speed_ms,0,blend_radius_m)
  movel([0.529262, -1.159941, -2.701744, -0.850704, 1.570796, 2.100059],accel_mss,speed_ms,0,blend_radius_m)
  speed_ms = 0.003
  movel([0.529262, -1.145084, -2.694241, -0.873064, 1.570796, 2.100059],accel_mss,speed_ms,0,blend_radius_m)
  speed_ms = 1.000
  movel([0.529262, -1.117192, -2.678884, -0.916313, 1.570796, 2.100059],accel_mss,speed_ms,0,blend_radius_m)
  movel([0.568778, -1.116819, -2.679036, -0.916534, 1.570796, 2.139574],accel_mss,speed_ms,0,blend_radius_m)
  movel([0.568778, -1.144712, -2.694398, -0.873279, 1.570796, 2.139574],accel_mss,speed_ms,0,blend_radius_m)
  speed_ms = 0.003
  movel([0.568778, -1.155797, -2.700039, -0.856554, 1.570796, 2.139574],accel_mss,speed_ms,0,blend_radius_m)
  speed_ms = 0.007
  movel([0.572935, -1.156054, -2.699928, -0.856406, 1.570796, 2.143731],accel_mss,speed_ms,0,blend_radius_m)
  movel([0.577080, -1.156333, -2.699809, -0.856247, 1.570796, 2.147877],accel_mss,speed_ms,0,blend_radius_m)
  movel([0.562608, -1.182829, -2.688096, -0.841464, 1.570796, 2.133405],accel_mss,speed_ms,0,blend_radius_m)
  movel([0.548864, -1.208191, -2.676183, -0.828015, 1.570796, 2.119661],accel_mss,speed_ms,0,blend_radius_m)
  movel([0.544954, -1.208238, -2.676160, -0.827991, 1.570796, 2.115751],accel_mss,speed_ms,0,blend_radius_m)
  movel([0.541035, -1.208305, -2.676128, -0.827957, 1.570796, 2.111831],accel_mss,speed_ms,0,blend_radius_m)
  movel([0.554543, -1.182631, -2.688186, -0.841572, 1.570796, 2.125340],accel_mss,speed_ms,0,blend_radius_m)
  movel([0.568778, -1.155797, -2.700039, -0.856554, 1.570796, 2.139574],accel_mss,speed_ms,0,blend_radius_m)
  speed_ms = 0.003
  movel([0.568778, -1.159570, -2.701904, -0.850916, 1.570796, 2.139574],accel_mss,speed_ms,0,blend_radius_m)
  speed_ms = 0.007
  movel([0.572935, -1.159827, -2.701793, -0.850769, 1.570796, 2.143731],accel_mss,speed_ms,0,blend_radius_m)
  movel([0.577080, -1.160105, -2.701673, -0.850611, 1.570796, 2.147877],accel_mss,speed_ms,0,blend_radius_m)
  movel([0.562608, -1.186571, -2.689915, -0.835903, 1.570796, 2.133405],accel_mss,speed_ms,0,blend_radius_m)
  movel([0.548864, -1.211898, -2.677959, -0.822532, 1.570796, 2.119661],accel_mss,speed_ms,0,blend_radius_m)
  movel([0.544954, -1.211945, -2.677936, -0.822508, 1.570796, 2.115751],accel_mss,speed_ms,0,blend_radius_m)
  movel([0.541035, -1.212012, -2.677903, -0.822474, 1.570796, 2.111831],accel_mss,speed_ms,0,blend_radius_m)
  movel([0.554543, -1.186374, -2.690005, -0.836010, 1.570796, 2.125340],accel_mss,speed_ms,0,blend_radius_m)
  movel([0.568778, -1.159570, -2.701904, -0.850916, 1.570796, 2.139574],accel_mss,speed_ms,0,blend_radius_m)
  speed_ms = 0.003
  movel([0.568778, -1.144712, -2.694398, -0.873279, 1.570796, 2.139574],accel_mss,speed_ms,0,blend_radius_m)
  speed_ms = 1.000
  movel([0.568778, -1.116819, -2.679036, -0.916534, 1.570796, 2.139574],accel_mss,speed_ms,0,blend_radius_m)
  movel([0.561419, -1.074141, -2.695584, -0.942664, 1.570796, 2.132216],accel_mss,speed_ms,0,blend_radius_m)
  movel([0.561419, -1.102092, -2.711496, -0.898802, 1.570796, 2.132216],accel_mss,speed_ms,0,blend_radius_m)
  speed_ms = 0.003
  movel([0.561419, -1.113247, -2.717349, -0.881793, 1.570796, 2.132216],accel_mss,speed_ms,0,blend_radius_m)
  speed_ms = 0.007
  movel([0.547356, -1.113009, -2.717441, -0.881939, 1.570796, 2.118152],accel_mss,speed_ms,0,blend_radius_m)
  movel([0.533169, -1.113014, -2.717439, -0.881936, 1.570796, 2.103966],accel_mss,speed_ms,0,blend_radius_m)
  movel([0.535280, -1.108714, -2.719091, -0.884584, 1.570796, 2.106077],accel_mss,speed_ms,0,blend_radius_m)
  movel([0.537409, -1.104383, -2.720737, -0.887269, 1.570796, 2.108205],accel_mss,speed_ms,0,blend_radius_m)
  movel([0.551697, -1.104377, -2.720739, -0.887272, 1.570796, 2.122493],accel_mss,speed_ms,0,blend_radius_m)
  movel([0.565859, -1.104621, -2.720647, -0.887121, 1.570796, 2.136655],accel_mss,speed_ms,0,blend_radius_m)
  movel([0.563630, -1.108949, -2.719001, -0.884439, 1.570796, 2.134426],accel_mss,speed_ms,0,blend_radius_m)
  movel([0.561419, -1.113247, -2.717349, -0.881793, 1.570796, 2.132216],accel_mss,speed_ms,0,blend_radius_m)
  speed_ms = 0.003
  movel([0.561419, -1.117051, -2.719285, -0.876053, 1.570796, 2.132216],accel_mss,speed_ms,0,blend_radius_m)
  speed_ms = 0.007
  movel([0.547356, -1.116813, -2.719378, -0.876199, 1.570796, 2.118152],accel_mss,speed_ms,0,blend_radius_m)
  movel([0.533169, -1.116818, -2.719376, -0.876196, 1.570796, 2.103966],accel_mss,speed_ms,0,blend_radius_m)
  movel([0.535280, -1.112519, -2.721035, -0.878835, 1.570796, 2.106077],accel_mss,speed_ms,0,blend_radius_m)
  movel([0.537409, -1.108189, -2.722688, -0.881511, 1.570796, 2.108205],accel_mss,speed_ms,0,blend_radius_m)
  movel([0.551697, -1.108184, -2.722690, -0.881514, 1.570796, 2.122493],accel_mss,speed_ms,0,blend_radius_m)
  movel([0.565859, -1.108427, -2.722598, -0.881364, 1.570796, 2.136655],accel_mss,speed_ms,0,blend_radius_m)
  movel([0.563630, -1.112754, -2.720944, -0.878690, 1.570796, 2.134426],accel_mss,speed_ms,0,blend_radius_m)
  movel([0.561419, -1.117051, -2.719285, -0.876053, 1.570796, 2.132216],accel_mss,speed_ms,0,blend_radius_m)
  speed_ms = 0.003
  movel([0.561419, -1.102092, -2.711496, -0.898802, 1.570796, 2.132216],accel_mss,speed_ms,0,blend_radius_m)
  speed_ms = 1.000
  movel([0.561419, -1.074141, -2.695584, -0.942664, 1.570796, 2.132216],accel_mss,speed_ms,0,blend_radius_m)
  movel([0.534542, -1.077420, -2.694371, -0.940598, 1.570796, 2.105338],accel_mss,speed_ms,0,blend_radius_m)
  movel([0.534542, -1.105372, -2.710241, -0.896776, 1.570796, 2.105338],accel_mss,speed_ms,0,blend_radius_m)
  speed_ms = 0.003
  movel([0.534542, -1.116525, -2.716077, -0.879787, 1.570796, 2.105338],accel_mss,speed_ms,0,blend_radius_m)
  speed_ms = 0.007
  movel([0.585441, -1.118073, -2.715474, -0.878843, 1.570796, 2.156237],accel_mss,speed_ms,0,blend_radius_m)
  movel([0.551443, -1.182164, -2.688399, -0.841826, 1.570796, 2.122239],accel_mss,speed_ms,0,blend_radius_m)
  movel([0.521341, -1.239997, -2.660224, -0.812167, 1.570796, 2.092138],accel_mss,speed_ms,0,blend_radius_m)
  movel([0.475369, -1.239016, -2.660734, -0.812639, 1.570796, 2.046166],accel_mss,speed_ms,0,blend_radius_m)
  movel([0.428294, -1.240385, -2.660022, -0.811981, 1.570796, 1.999090],accel_mss,speed_ms,0,blend_radius_m)
  movel([0.453497, -1.182431, -2.688277, -0.841681, 1.570796, 2.024293],accel_mss,speed_ms,0,blend_radius_m)
  movel([0.482054, -1.118193, -2.715427, -0.878770, 1.570796, 2.052850],accel_mss,speed_ms,0,blend_radius_m)
  movel([0.534542, -1.116525, -2.716077, -0.879787, 1.570796, 2.105338],accel_mss,speed_ms,0,blend_radius_m)
  speed_ms = 0.003
  movel([0.534542, -1.120327, -2.718009, -0.874054, 1.570796, 2.105338],accel_mss,speed_ms,0,blend_radius_m)
  speed_ms = 0.007
  movel([0.585441, -1.121873, -2.717402, -0.873113, 1.570796, 2.156237],accel_mss,speed_ms,0,blend_radius_m)
  movel([0.551443, -1.185908, -2.690219, -0.836262, 1.570796, 2.122239],accel_mss,speed_ms,0,blend_radius_m)
  movel([0.521341, -1.243652, -2.661945, -0.806792, 1.570796, 2.092138],accel_mss,speed_ms,0,blend_radius_m)
  movel([0.475369, -1.242672, -2.662457, -0.807260, 1.570796, 2.046166],accel_mss,speed_ms,0,blend_radius_m)
  movel([0.428294, -1.244039, -2.661742, -0.806607, 1.570796, 1.999090],accel_mss,speed_ms,0,blend_radius_m)
  movel([0.453497, -1.186174, -2.690097, -0.836118, 1.570796, 2.024293],accel_mss,speed_ms,0,blend_radius_m)
  movel([0.482054, -1.121993, -2.717355, -0.873041, 1.570796, 2.052850],accel_mss,speed_ms,0,blend_radius_m)
  movel([0.534542, -1.120327, -2.718009, -0.874054, 1.570796, 2.105338],accel_mss,speed_ms,0,blend_radius_m)
  speed_ms = 0.003
  movel([0.534542, -1.105372, -2.710241, -0.896776, 1.570796, 2.105338],accel_mss,speed_ms,0,blend_radius_m)
  speed_ms = 1.000
  movel([0.534542, -1.077420, -2.694371, -0.940598, 1.570796, 2.105338],accel_mss,speed_ms,0,blend_radius_m)
  movel([0.061043, -1.173967, -2.654157, -0.884264, 1.570796, 1.631840],accel_mss,speed_ms,0,blend_radius_m)
  movel([0.061043, -1.080275, -2.588658, -1.043456, 1.570796, 1.631840],accel_mss,speed_ms,0,blend_radius_m)
  # End of main program
